{region 'Documentation'}
(*!
<summary>Checks that IN is positive or negative infinity.</summary>
<description>

NaN and either infinity are legitimate checked data, not configuration errors.
Classification mismatch reports Failed. Bit-based classification does not perform an ordered
floating-point comparison.

Numeric diagnostics use the formatter's default six significant digits; rounding affects
the message only, not the comparison.

</description>
*)
{endregion}
FUNCTION_BLOCK AssertIsInfinite_LReal EXTENDS AssertionBase
VAR_INPUT
    IN : LREAL; //! Value to classify; NaN and both infinities are valid inputs.
END_VAR

SUPER^();

{region 'Documentation'}
(*!
<summary>Classifies the bit representation without floating-point arithmetic.</summary>
*)
{endregion}
METHOD PROTECTED Assert
VAR
    Representation : AssertionLRealRepresentation;
    Message : STRING(GVL_Constants.MessageLength);
END_VAR
VAR CONSTANT
    ExponentMask : LWORD := LWORD#16#7FF0000000000000;
    FractionMask : LWORD := LWORD#16#000FFFFFFFFFFFFF;
END_VAR
IF NOT EvaluationActive THEN
    RETURN;
END_IF;

IF Result = E_Result.Error THEN
    RETURN;
END_IF;

IF Result = E_Result.Failed THEN
    RETURN;
END_IF;

Representation.Value := IN;
IF ((Representation.Bits AND ExponentMask) <> ExponentMask)
    OR ((Representation.Bits AND FractionMask) <> 0) THEN
    Message := CONCAT('Assertion failed: expected positive or negative infinity. Actual = ',
        CreateAssertionTextValue_LReal(Value := IN));
    Message := CONCAT(Message, '.');
    Fail(Message := Message);
    RETURN;
END_IF;

Pass();
END_METHOD

END_FUNCTION_BLOCK

(* stored: Version 1.1.0.1
   POU AssertIsInfinite_LReal: Id {fe969339-6314-4876-b1a4-a6906c5f4868}, SpecialFunc None
   Folder Internal: Id {4ef9a8df-49bd-4d80-a97f-a52cc43db226}
   Method Assert: Id {a6310000-0000-4000-8000-000000000005} *)
